SUBAPPLICATION FU_Sollwert (* Sollfrequenz in Hz vom Web-Dashboard (OPC UA FU1.SollFrequenz) -> auf 0..Fmax begrenzen -> % von Fmax -> 9301H. *)
  (* Standard: 61499-2; Description: Copyright (c) 2026 Franz Höpfinger This program and the accompanying materials are made available under the terms of the Eclipse Public License 2.0 which is available at https://www.eclipse.org/legal/epl-2.0/ SPDX-License-Identifier: EPL-2.0 *)
  (* Version 1.0, 2026-11-02, Franz Höpfinger, Franz Höpfinger, aus FU_Demo_H300 herausgeloest *)
  PACKAGE FBs::FU_Demo;
  IMPORT FBs::FU_Demo::FU_Demo_Konstanten::FU_MODBUS_SOLLWERT;
  IMPORT FBs::FU_Demo::FU_Demo_Konstanten::FU_FMAX_HZ;
  IMPORT FBs::FU_Demo::FU_Demo_Konstanten::FU_SOLLWERT_FAKTOR;
  IMPORT FBs::FU_Demo::FU_Demo_Konstanten::FU_SOLLFREQUENZ_WEB_READ;
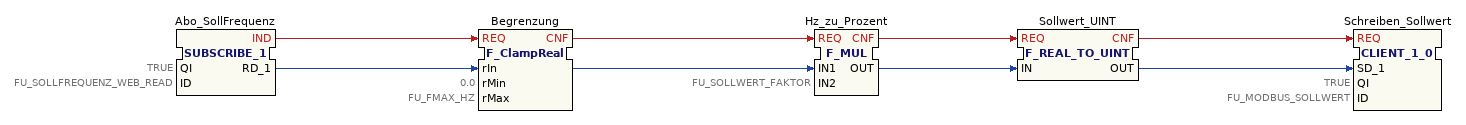
  FBS
    Abo_SollFrequenz : iec61499::net::SUBSCRIBE_1(QI := TRUE, ID := FU_SOLLFREQUENZ_WEB_READ);
    Begrenzung : logiBUS::signalprocessing::clamp::F_ClampReal(rMin := 0.0, rMax := FU_FMAX_HZ); (* 0 .. Fmax Hz; typisiert den OPC-UA-Knoten als Float *)
    Hz_zu_Prozent : iec61131::arithmetic::F_MUL(IN2 := FU_SOLLWERT_FAKTOR); (* Hz * 10000 / Fmax = Registerwert 9301H (0..10000) *)
    Sollwert_UINT : iec61131::conversion::F_REAL_TO_UINT;
    Schreiben_Sollwert : iec61499::net::CLIENT_1_0(QI := TRUE, ID := FU_MODBUS_SOLLWERT); (* 9301H Frequenzsollwert *)
  END_FBS
  EVENT_CONNECTIONS
    Abo_SollFrequenz.IND TO Begrenzung.REQ;
    Begrenzung.CNF TO Hz_zu_Prozent.REQ;
    Hz_zu_Prozent.CNF TO Sollwert_UINT.REQ;
    Sollwert_UINT.CNF TO Schreiben_Sollwert.REQ;
  END_CONNECTIONS
  DATA_CONNECTIONS
    Abo_SollFrequenz.RD_1 TO Begrenzung.rIn;
    Begrenzung. TO Hz_zu_Prozent.IN1;
    Hz_zu_Prozent.OUT TO Sollwert_UINT.IN;
    Sollwert_UINT.OUT TO Schreiben_Sollwert.SD_1;
  END_CONNECTIONS
END_SUBAPPLICATION
